(*
SPDX-FileCopyrightText: c 2026 Oleksandr Tiutyk <trofimich@gmail.com>
SPDX-License-Identifier: MIT
License: https://opensource.org/license/mit
*)

(*!
<summary>Groups wide-string formatting, editing, search and splitter contracts.</summary>
<description>
Owns the independent child instances and their fixed registration array. Use from one PLC task at a stable address.
</description>
*)

{attribute 'no_assign'}
{attribute 'no_explicit_call' := 'do not call this function block directly'}
FUNCTION_BLOCK WideStringsTestGroup EXTENDS TOF_Testing.TestGroup<11>
VAR_STAT
	{attribute 'hide'}
	_ClassName : STRING := __POUNAME();
END_VAR
VAR
	_AnyToStringFit255 : WideStringFitFormattingTest(name := "AnyToStringFit255", parent := THIS^);
	_Append : WideStringAppendTest(name := "Append", parent := THIS^);
	_AppendFit : WideStringAppendFitTest(name := "AppendFit", parent := THIS^);
	_ConcatFit255 : WideStringConcatFitTest(name := "ConcatFit255", parent := THIS^);
	_Contains : WideStringContainsTest(name := "Contains", parent := THIS^);
	_Join : WideStringJoinTest(name := "Join", parent := THIS^);
	_ReplaceInSource : WideStringReplacementTest(name := "ReplaceInSource", parent := THIS^);
	_Split : WideStringSplitTest(name := "Split", parent := THIS^);
	_Trim : WideStringTrimTest(name := "Trim", parent := THIS^);
	_SplitterSeparatorBounds : WideStringSeparatorBoundsTest(name := "SplitterSeparatorBounds", parent := THIS^);
	_AnyToStringFitLongInputs : WideStringLongFitFormattingTest(name := "AnyToStringFitLongInputs", parent := THIS^);

	_Children : ARRAY [0.._ChildCount - 1] OF TOF_Testing.ITestElement :=
	[
		_AnyToStringFit255,
		_Append,
		_AppendFit,
		_ConcatFit255,
		_Contains,
		_Join,
		_ReplaceInSource,
		_Split,
		_Trim,
		_SplitterSeparatorBounds,
		_AnyToStringFitLongInputs
	];
END_VAR

//! <summary>Borrows the fixed child array. Callers must not modify it.</summary>
{attribute 'monitoring' := 'call'}
PROPERTY Children : REFERENCE TO ARRAY [0.._ChildCount - 1] OF TOF_Testing.ITestElement
GET
Children REF= _Children;
END_GET
END_PROPERTY

//! <summary>Borrows the concrete class name. Callers must not modify it.</summary>
{attribute 'monitoring' := 'call'}
PROPERTY ClassName : REFERENCE TO STRING
GET
ClassName REF= _ClassName;
END_GET
END_PROPERTY

//! <summary>Borrows the compiler-initialized namespace name. Callers must not modify it.</summary>
{attribute 'monitoring' := 'call'}
PROPERTY NamespaceName : REFERENCE TO STRING
GET
NamespaceName REF= CurrentNamespace.Name;
END_GET
END_PROPERTY

//! <summary>Reports the concrete instance size in bytes.</summary>
{attribute 'monitoring' := 'call'}
PROPERTY SelfSize : ULINT
GET
SelfSize := XSIZEOF(THIS^);
END_GET
END_PROPERTY

END_FUNCTION_BLOCK

(* stored: Version 1.1.0.1
   POU WideStringsTestGroup: Id {edc3fc4a-c574-4eed-93db-6d5af7501ae4}, SpecialFunc None
   Property Children: Id {88f66cc8-dc2a-4b1c-bfc3-b7a0d84f963a}
   Get Get: Id {d532122e-6655-437a-aa30-f526366bcb11}
   Property ClassName: Id {5e728a1a-73b0-4356-ad10-6319e34c2081}
   Get Get: Id {10d294dd-2858-45cb-a0bb-0aa95b7920b4}
   Property NamespaceName: Id {50e83767-8d50-4bd5-bb2d-9b88013405a3}
   Get Get: Id {9a000aaf-e4b2-434d-8f51-c2c50288ad2c}
   Property SelfSize: Id {71de2408-7c69-4beb-a2a8-2653711be038}
   Get Get: Id {622d0643-3993-4ba4-9f87-b3a2cb118713} *)
